(* IEC 61131-3 sources: llm-plc-st-eval/data/definitivo/gpt-4o-2024-08-06/I1/few_shot, 3 files *)

(* ---- ejec_1.st ---- *)
```pascal
FUNCTION_BLOCK FB_Semaforo
VAR_INPUT
    habilitado : BOOL; (* Habilitacion del semaforo *)
END_VAR
VAR_OUTPUT
    luzV : BOOL; (* Luz verde *)
    luzA : BOOL; (* Luz amarilla *)
    luzR : BOOL; (* Luz roja *)
END_VAR
VAR
    tCiclo : TON; (* Temporizador para el ciclo del semaforo *)
    tIntermitente : TON; (* Temporizador para el amarillo intermitente *)
    estado : INT; (* Estado del semaforo *)
    intermitente : BOOL; (* Estado de la luz amarilla intermitente *)
END_VAR

(* Logica del semaforo *)
IF habilitado THEN
    (* Control del ciclo del semaforo *)
    CASE estado OF
        0: (* Luz verde *)
            luzV := TRUE;
            luzA := FALSE;
            luzR := FALSE;
            tCiclo(IN := TRUE, PT := T#20S);
            IF tCiclo.Q THEN
                estado := 1;
                tCiclo(IN := FALSE);
            END_IF;
        1: (* Luz amarilla *)
            luzV := FALSE;
            luzA := TRUE;
            luzR := FALSE;
            tCiclo(IN := TRUE, PT := T#4S);
            IF tCiclo.Q THEN
                estado := 2;
                tCiclo(IN := FALSE);
            END_IF;
        2: (* Luz roja *)
            luzV := FALSE;
            luzA := FALSE;
            luzR := TRUE;
            tCiclo(IN := TRUE, PT := T#15S);
            IF tCiclo.Q THEN
                estado := 0;
                tCiclo(IN := FALSE);
            END_IF;
    END_CASE;
ELSE
    (* Control del amarillo intermitente *)
    luzV := FALSE;
    luzR := FALSE;
    tIntermitente(IN := TRUE, PT := T#1S);
    IF tIntermitente.Q THEN
        intermitente := NOT intermitente;
        tIntermitente(IN := FALSE);
    END_IF;
    luzA := intermitente;
    estado := 0; (* Reiniciar ciclo al habilitar *)
END_IF;
END_FUNCTION_BLOCK
```

(* ---- ejec_2.st ---- *)
```pascal
FUNCTION_BLOCK FB_Semaforo
VAR_INPUT
    habilitado : BOOL; (* Habilitacion del semaforo *)
END_VAR
VAR_OUTPUT
    luzV : BOOL; (* Luz verde *)
    luzA : BOOL; (* Luz amarilla *)
    luzR : BOOL; (* Luz roja *)
END_VAR
VAR
    tCiclo : TON; (* Temporizador para el ciclo del semaforo *)
    tIntermitente : TON; (* Temporizador para el amarillo intermitente *)
    estado : INT; (* Estado del semaforo *)
END_VAR

(* Inicializacion de variables *)
IF NOT habilitado THEN
    (* Modo amarillo intermitente *)
    tIntermitente(IN := TRUE, PT := T#1S);
    luzV := FALSE;
    luzR := FALSE;
    luzA := tIntermitente.Q;
    tCiclo(IN := FALSE);
    estado := 0; (* Reiniciar estado al habilitar de nuevo *)
ELSE
    (* Modo ciclo normal del semaforo *)
    tIntermitente(IN := FALSE);
    CASE estado OF
        0: (* Luz verde *)
            luzV := TRUE;
            luzA := FALSE;
            luzR := FALSE;
            tCiclo(IN := TRUE, PT := T#20S);
            IF tCiclo.Q THEN
                estado := 1;
                tCiclo(IN := FALSE);
            END_IF
        1: (* Luz amarilla *)
            luzV := FALSE;
            luzA := TRUE;
            luzR := FALSE;
            tCiclo(IN := TRUE, PT := T#4S);
            IF tCiclo.Q THEN
                estado := 2;
                tCiclo(IN := FALSE);
            END_IF
        2: (* Luz roja *)
            luzV := FALSE;
            luzA := FALSE;
            luzR := TRUE;
            tCiclo(IN := TRUE, PT := T#15S);
            IF tCiclo.Q THEN
                estado := 0;
                tCiclo(IN := FALSE);
            END_IF
    END_CASE
END_IF
END_FUNCTION_BLOCK
```

(* ---- ejec_3.st ---- *)
```pascal
FUNCTION_BLOCK FB_Semaforo
VAR_INPUT
    habilitado : BOOL; (* Habilitacion del semaforo *)
END_VAR
VAR_OUTPUT
    luzV : BOOL; (* Luz verde *)
    luzA : BOOL; (* Luz amarilla *)
    luzR : BOOL; (* Luz roja *)
END_VAR
VAR
    tCiclo : TON; (* Temporizador para el ciclo del semaforo *)
    tIntermitente : TON; (* Temporizador para el amarillo intermitente *)
    estado : INT; (* Estado del semaforo *)
    intermitente : BOOL; (* Estado del intermitente *)
END_VAR

(* Logica del semaforo ciclico *)
IF habilitado THEN
    (* Control del ciclo del semaforo *)
    CASE estado OF
        0: (* Verde 20 segundos *)
            luzV := TRUE;
            luzA := FALSE;
            luzR := FALSE;
            tCiclo(IN := TRUE, PT := T#20S);
            IF tCiclo.Q THEN
                estado := 1;
                tCiclo(IN := FALSE);
            END_IF;
        1: (* Amarillo 4 segundos *)
            luzV := FALSE;
            luzA := TRUE;
            luzR := FALSE;
            tCiclo(IN := TRUE, PT := T#4S);
            IF tCiclo.Q THEN
                estado := 2;
                tCiclo(IN := FALSE);
            END_IF;
        2: (* Rojo 15 segundos *)
            luzV := FALSE;
            luzA := FALSE;
            luzR := TRUE;
            tCiclo(IN := TRUE, PT := T#15S);
            IF tCiclo.Q THEN
                estado := 0;
                tCiclo(IN := FALSE);
            END_IF;
    END_CASE;
ELSE
    (* Amarillo intermitente *)
    luzV := FALSE;
    luzR := FALSE;
    tIntermitente(IN := TRUE, PT := T#1S);
    IF tIntermitente.Q THEN
        intermitente := NOT intermitente;
        tIntermitente(IN := FALSE);
    END_IF;
    luzA := intermitente;
    estado := 0; (* Reinicia el ciclo al habilitar *)
END_IF;
END_FUNCTION_BLOCK
```
